{attribute 'qualified_only'}
//{attribute 'strict'}
{attribute 'to_string'}
TYPE E_Element_List :
(
eNotSelected := 0,
eTank_1,
eTank_2,
eTank_3,
eTank_4,
eTriBlender_Marinada,
eTriBlender_Color,
eLine_Marinada,
eLine_Color
);
END_TYPE

(* stored: Version 1.1.0.1, ProductVersion 3.1.4024.12
   DUT E_Element_List: Id {5307231e-88b6-4a18-8b65-faf2eefebe7f} *)
